Fanuc KAREL source: kt00519.KL

-- PROVISIONAL review KL for V940-1; original PC SHA256 1dc8353bff4e44fbbf6cbafaef3bb9f4b662e13f497f4b086c4dfa4f08e67694
-- Incomplete behavior may be omitted. Consult companion uncertainty JSON. Do not deploy.
PROGRAM KT00519
%NOLOCKGROUP
-- UNRESOLVED_DECL P1 type=000106
-- UNRESOLVED_DECL P2 type=000102
-- UNRESOLVED_DECL OUT type=000101
BEGIN
  -- V9_ZERO_TABLE_METADATA_HINT layout=0001; no indexed target words; source/name/runtime held
  -- UNRESOLVED_PC offsets 5-20; opcodes 2E,22,32,35
  -- UNRESOLVED_PC offsets 25-40; opcodes 2E,22,32,35
  -- UNRESOLVED_PC offsets 45-79; opcodes 49,7E,49,7E,60,4A
  -- UNRESOLVED_PC offsets 84-88; opcodes 7F
END KT00519
